Fanuc KAREL source: kt00133.KL

-- PROVISIONAL review KL for V770-1; original PC SHA256 54e78fc9e3118907bd2599bf0c7e0938885214c7294d6ab4e35dd820a31cc649
-- Incomplete behavior may be omitted. Consult companion uncertainty JSON. Do not deploy.
PROGRAM KT00133
%NOLOCKGROUP
VAR
  I1 : INTEGER
  OUT : INTEGER
-- UNRESOLVED_DECL Y2 type=002018
BEGIN
  -- UNRESOLVED_PC offsets 5-16; opcodes 2E,23
  -- UNRESOLVED_PC offsets 21-35; opcodes 2E,22,9D,33,B2
  -- UNRESOLVED_PC offsets 40-62; opcodes 21,22,9D,33,B1,55,23
  -- UNRESOLVED_PC offsets 67-71; opcodes 7F
END KT00133
